// TIA Portal V20 export
VAR_GLOBAL   // PLC tag table "LASER_OUT_datalogic"
   START_MARKING AT %Q1500.0 : Bool;
   STOP_SYSTEM AT %Q1500.1 : Bool;
   GET_PNIO_PROTOCOL_VERSION AT %Q1501.0 : Bool;
   PROTOCOL_ERROR_CLEAR AT %Q1501.7 : Bool;
   OPEN_DOKUMENT_FROM_DEVICE AT %Q1502.0 : Bool;
   SAVE_DOKUMENT AT %Q1502.1 : Bool;
   GET_DATA_FIELD_VALUE AT %Q1502.2 : Bool;
   SET_DATA_FIELD_VALUE AT %Q1502.3 : Bool;
   GET_GLOBAL_COUNTER_VALUE AT %Q1502.4 : Bool;
   SET_GLOBAL_COUNTER_VALUE AT %Q1502.5 : Bool;
   GET_GLOBAL_STRING_VALUE AT %Q1502.6 : Bool;
   SET_GLOBAL_STRING_VALUE AT %Q1502.7 : Bool;
   ENABLE_DATA_FIELD AT %Q1503.0 : Bool;
   DISABLE_DATA_FIELD AT %Q1503.1 : Bool;
   MOVE_AND_ROTATE_DOCUMENT AT %Q1504.0 : Bool;
   MOVE_DATA_FIELD AT %Q1504.1 : Bool;
   RESERVE_Q_5_BYTE AT %QB1505 : Byte;
   RESERVE_Q_6_BYTE AT %QB1506 : Byte;
   RESERVE_Q_7_BYTE AT %QB1507 : Byte;
   MOVE_AXIS AT %Q1508.0 : Bool;
   RESET_AXIS AT %Q1508.1 : Bool;
   STOP_AXIS AT %Q1508.2 : Bool;
   START_AUTOFOCUS AT %Q1508.3 : Bool;
   STOP_AUTOFOCUS AT %Q1508.4 : Bool;
   SET_FOCUS_DISTANCE_SENSOR_REFERENCE AT %Q1508.5 : Bool;
   RESERVE_Q_9_BYTE AT %QB1509 : Byte;
   X_AXIS AT %Q1510.0 : Bool;
   Y_AXIS AT %Q1510.1 : Bool;
   Z_AXIS AT %Q1510.2 : Bool;
   R_AXIS AT %Q1510.3 : Bool;
   RESERVE_Q_11_BYTE AT %QB411 : Byte;
   RESERVE_Q_12_BYTE AT %QB412 : Byte;
   RESERVE_Q_13_BYTE AT %QB413 : Byte;
   RESERVE_Q_14_BYTE AT %QB414 : Byte;
   RESERVE_Q_15_BYTE AT %QB415 : Byte;
   RESERVE_Q_16_BYTE AT %QB416 : Byte;
   RESERVE_Q_17_BYTE AT %QB417 : Byte;
   RESERVE_Q_18_BYTE AT %QB418 : Byte;
   RESERVE_Q_19_BYTE AT %QB419 : Byte;
   RESERVE_Q_20_BYTE AT %QB420 : Byte;
   RESERVE_Q_21_BYTE AT %QB421 : Byte;
   SET_AUTPUT AT %Q1522.0 : Bool;
   RESET_OUTPUT AT %Q1522.1 : Bool;
   RESERVE_Q_23_BYTE AT %QB1523 : Byte;   // --------------------
   I_O_PORT_LASER_OUTPUT_0 AT %Q1524.0 : Bool;
   I_O_PORT_LASER_OUTPUT_1 AT %Q1524.1 : Bool;
   I_O_PORT_LASER_OUTPUT_2 AT %Q1524.2 : Bool;
   I_O_PORT_LASER_OUTPUT_3 AT %Q1524.3 : Bool;
   I_O_PORT_LASER_OUTPUT_4 AT %Q1524.4 : Bool;
   I_O_PORT_LASER_OUTPUT_5 AT %Q1524.5 : Bool;
   I_O_PORT_LASER_OUTPUT_6 AT %Q1524.6 : Bool;
   I_O_PORT_LASER_OUTPUT_7 AT %Q1524.7 : Bool;
   I_O_PORT_LASER_OUTPUT_8 AT %Q1525.0 : Bool;
   I_O_PORT_LASER_OUTPUT_9 AT %Q1525.1 : Bool;
   I_O_PORT_LASER_OUTPUT_10 AT %Q1525.2 : Bool;
   I_O_PORT_LASER_OUTPUT_11 AT %Q1525.3 : Bool;
   I_O_PORT_LASER_OUTPUT_12 AT %Q1525.4 : Bool;
   I_O_PORT_LASER_OUTPUT_13 AT %Q1525.5 : Bool;
   I_O_PORT_LASER_OUTPUT_14 AT %Q1525.6 : Bool;
   I_O_PORT_LASER_OUTPUT_15 AT %Q1525.7 : Bool;
   RESERVE_Q_26_BYTE AT %QB1526 : Byte;   // --------------------
   RESERVE_Q_27_BYTE AT %QB1527 : Byte;   // --------------------
   RESERVE_Q_28_BYTE AT %QB1528 : Byte;   // --------------------
   RESERVE_Q_29_BYTE AT %QB1529 : Byte;   // --------------------
   RESERVE_Q_30_BYTE AT %QB1530 : Byte;   // --------------------
   RESERVE_Q_31_BYTE AT %QB1531 : Byte;   // --------------------
   GET_ID_MATCH_RESULT AT %Q1532.1 : Bool;
   GET_ID_MARVIS_CONFIGURATION AT %Q1532.2 : Bool;
   SET_ID_MARVIS_CONFIGURATION AT %Q1532.3 : Bool;
   GET_ID_MARVIS_RESULT AT %Q1532.4 : Bool;
   RESERVE_Q_33_BYTE AT %QB1533 : Byte;
   RESERVE_Q_34_BYTE AT %QB1534 : Byte;
   RESERVE_Q_35_BYTE AT %QB1535 : Byte;
   RESERVE_Q_36_BYTE AT %QB1536 : Byte;
   RESERVE_Q_37_BYTE AT %QB1537 : Byte;
   RESERVE_Q_38_BYTE AT %QB1538 : Byte;
   RESERVE_Q_39_BYTE AT %QB1539 : Byte;
   RESERVE_Q_40_BYTE AT %QB1540 : Byte;
   RESERVE_Q_41_BYTE AT %QB1541 : Byte;
   RESERVE_Q_42_BYTE AT %QB1542 : Byte;
   RESERVE_Q_43_BYTE AT %QB1543 : Byte;
   RESERVE_Q_44_BYTE AT %QB1544 : Byte;
   RESERVE_Q_45_BYTE AT %QB1545 : Byte;
   RESERVE_Q_46_BYTE AT %QB1546 : Byte;
   RESERVE_Q_47_BYTE AT %QB1547 : Byte;
   RESERVE_Q_48_BYTE AT %QB1548 : Byte;
   RESERVE_Q_49_BYTE AT %QB1549 : Byte;
   RESERVE_Q_50_BYTE AT %QB1550 : Byte;
   RESERVE_Q_51_BYTE AT %QB1551 : Byte;
   RESERVE_Q_52_BYTE AT %QB1552 : Byte;
   RESERVE_Q_53_BYTE AT %QB1553 : Byte;
   REQUEST_DATA_SIZE AT %QB1554 : Byte;
   RESERVE_Q_55_BYTE AT %QB1555 : Byte;
   REQUEST_DATA_FIELC_BYTE_0 AT %QB1556 : Byte;
   REQUEST_DATA_FIELC_BYTE_1 AT %QB1557 : Byte;
   REQUEST_DATA_FIELC_BYTE_2 AT %QB1558 : Byte;
   REQUEST_DATA_FIELC_BYTE_3 AT %QB1559 : Byte;
   REQUEST_DATA_FIELC_BYTE_4 AT %QB1560 : Byte;
   REQUEST_DATA_FIELC_BYTE_5 AT %QB1561 : Byte;
   REQUEST_DATA_FIELC_BYTE_6 AT %QB1562 : Byte;
   REQUEST_DATA_FIELC_BYTE_7 AT %QB1563 : Byte;
   REQUEST_DATA_FIELC_BYTE_8 AT %QB1564 : Byte;
   REQUEST_DATA_FIELC_BYTE_9 AT %QB1565 : Byte;
   REQUEST_DATA_FIELC_BYTE_10 AT %QB1566 : Byte;
   REQUEST_DATA_FIELC_BYTE_11 AT %QB1567 : Byte;
   REQUEST_DATA_FIELC_BYTE_12 AT %QB1568 : Byte;
   REQUEST_DATA_FIELC_BYTE_13 AT %QB1569 : Byte;
   REQUEST_DATA_FIELC_BYTE_14 AT %QB1570 : Byte;
   REQUEST_DATA_FIELC_BYTE_15 AT %QB1571 : Byte;
   REQUEST_DATA_FIELC_BYTE_16 AT %QB1572 : Byte;
   REQUEST_DATA_FIELC_BYTE_17 AT %QB1573 : Byte;
   REQUEST_DATA_FIELC_BYTE_18 AT %QB1574 : Byte;
   REQUEST_DATA_FIELC_BYTE_19 AT %QB1575 : Byte;
   REQUEST_DATA_FIELC_BYTE_20 AT %QB1576 : Byte;
   REQUEST_DATA_FIELC_BYTE_21 AT %QB1577 : Byte;
   REQUEST_DATA_FIELC_BYTE_22 AT %QB1578 : Byte;
   REQUEST_DATA_FIELC_BYTE_23 AT %QB1579 : Byte;
   REQUEST_DATA_FIELC_BYTE_24 AT %QB1580 : Byte;
   REQUEST_DATA_FIELC_BYTE_25 AT %QB1581 : Byte;
   REQUEST_DATA_FIELC_BYTE_26 AT %QB1582 : Byte;
   REQUEST_DATA_FIELC_BYTE_27 AT %QB1583 : Byte;
   REQUEST_DATA_FIELC_BYTE_28 AT %QB1584 : Byte;
   REQUEST_DATA_FIELC_BYTE_29 AT %QB1585 : Byte;
   REQUEST_DATA_FIELC_BYTE_30 AT %QB1586 : Byte;
   REQUEST_DATA_FIELC_BYTE_31 AT %QB1587 : Byte;
   REQUEST_DATA_FIELC_BYTE_32 AT %QB1588 : Byte;
   REQUEST_DATA_FIELC_BYTE_33 AT %QB1589 : Byte;
   REQUEST_DATA_FIELC_BYTE_34 AT %QB1590 : Byte;
   REQUEST_DATA_FIELC_BYTE_35 AT %QB1591 : Byte;
   REQUEST_DATA_FIELC_BYTE_36 AT %QB1592 : Byte;
   REQUEST_DATA_FIELC_BYTE_37 AT %QB1593 : Byte;
   REQUEST_DATA_FIELC_BYTE_38 AT %QB1594 : Byte;
   REQUEST_DATA_FIELC_BYTE_39 AT %QB1595 : Byte;
   REQUEST_DATA_FIELC_BYTE_40 AT %QB1596 : Byte;
   REQUEST_DATA_FIELC_BYTE_41 AT %QB1597 : Byte;
   REQUEST_DATA_FIELC_BYTE_42 AT %QB1598 : Byte;
   REQUEST_DATA_FIELC_BYTE_43 AT %QB1599 : Byte;
   REQUEST_DATA_FIELC_BYTE_44 AT %QB1600 : Byte;
   REQUEST_DATA_FIELC_BYTE_45 AT %QB1601 : Byte;
   REQUEST_DATA_FIELC_BYTE_46 AT %QB1602 : Byte;
   REQUEST_DATA_FIELC_BYTE_47 AT %QB1603 : Byte;
   REQUEST_DATA_FIELC_BYTE_48 AT %QB1604 : Byte;
   REQUEST_DATA_FIELC_BYTE_49 AT %QB1605 : Byte;
   REQUEST_DATA_FIELC_BYTE_50 AT %QB1606 : Byte;
   REQUEST_DATA_FIELC_BYTE_51 AT %QB1607 : Byte;
   REQUEST_DATA_FIELC_BYTE_52 AT %QB1608 : Byte;
   REQUEST_DATA_FIELC_BYTE_53 AT %QB1609 : Byte;
   REQUEST_DATA_FIELC_BYTE_54 AT %QB1610 : Byte;
   REQUEST_DATA_FIELC_BYTE_55 AT %QB1611 : Byte;
   REQUEST_DATA_FIELC_BYTE_56 AT %QB1612 : Byte;
   REQUEST_DATA_FIELC_BYTE_57 AT %QB1613 : Byte;
   REQUEST_DATA_FIELC_BYTE_58 AT %QB1614 : Byte;
   REQUEST_DATA_FIELC_BYTE_59 AT %QB1615 : Byte;
   REQUEST_DATA_FIELC_BYTE_60 AT %QB1616 : Byte;
   REQUEST_DATA_FIELC_BYTE_61 AT %QB1617 : Byte;
   REQUEST_DATA_FIELC_BYTE_62 AT %QB1618 : Byte;
   REQUEST_DATA_FIELC_BYTE_63 AT %QB1619 : Byte;
   REQUEST_DATA_FIELC_BYTE_64 AT %QB1620 : Byte;
   REQUEST_DATA_FIELC_BYTE_65 AT %QB1621 : Byte;
   REQUEST_DATA_FIELC_BYTE_66 AT %QB1622 : Byte;
   REQUEST_DATA_FIELC_BYTE_67 AT %QB1623 : Byte;
   REQUEST_DATA_FIELC_BYTE_68 AT %QB1624 : Byte;
   REQUEST_DATA_FIELC_BYTE_69 AT %QB1625 : Byte;
   REQUEST_DATA_FIELC_BYTE_70 AT %QB1626 : Byte;
   REQUEST_DATA_FIELC_BYTE_71 AT %QB1627 : Byte;
END_VAR
